(* IEC 61131-3 sources: trust-platform/examples/OSCAT/production_queue/non-oop/src, 3 files *)

(* ---- Configuration.st ---- *)
CONFIGURATION ProductionQueueClassicConfiguration
RESOURCE Cpu0 ON PLC
    TASK MainTask (INTERVAL := T#100ms, PRIORITY := 1);
    PROGRAM Main WITH MainTask : Main;
END_RESOURCE
END_CONFIGURATION

(* ---- Main.st ---- *)
PROGRAM Main
VAR
    OrderQueue : FIFO_16;
    NextOrderId : DWORD;
    QueueEmpty : BOOL;
END_VAR

OrderQueue(DIN := DWORD#16#1001, E := TRUE, RD := FALSE, WD := TRUE, RST := FALSE);
OrderQueue(DIN := DWORD#0, E := TRUE, RD := TRUE, WD := FALSE, RST := FALSE);
NextOrderId := OrderQueue.DOUT;
QueueEmpty := OrderQueue.EMPTY;
END_PROGRAM

(* ---- Tests.st ---- *)
TEST_PROGRAM ProductionQueueClassicPushesAndPopsOrderId
VAR
    OrderQueue : FIFO_16;
END_VAR

OrderQueue(DIN := DWORD#0, E := TRUE, RD := FALSE, WD := FALSE, RST := TRUE);
OrderQueue(DIN := DWORD#16#1001, E := TRUE, RD := FALSE, WD := TRUE, RST := FALSE);
OrderQueue(DIN := DWORD#0, E := TRUE, RD := TRUE, WD := FALSE, RST := FALSE);

ASSERT_EQUAL(EXPECTED := DWORD#16#1001, ACTUAL := OrderQueue.DOUT);
ASSERT_TRUE(IN := OrderQueue.EMPTY);
END_TEST_PROGRAM
